Fanuc KAREL source: CA0036.KL

PROGRAM CA0036
%STACKSIZE=65535
%PRIORITY=65535
%NOLOCKGROUP
TYPE
T=STRUCTURE
A : INTEGER
B : REAL
ENDSTRUCTURE
VAR
G : INTEGER
I : INTEGER
R : REAL
B : BOOLEAN
S : STRING[16]
AI : ARRAY[2] OF INTEGER
AR : ARRAY[2] OF REAL
ST : T
P : XYZWPR
V : VECTOR
ROUTINE F(P1 : ARRAY[*] OF INTEGER; P2 : ARRAY[*] OF REAL; P3 : T; P4 : XYZWPR; P5 : VECTOR; P6 : ARRAY[*] OF INTEGER; P7 : ARRAY[*] OF REAL; P8 : T; P9 : XYZWPR; P10 : VECTOR; P11 : ARRAY[*] OF INTEGER;
P12 : ARRAY[*] OF REAL) FROM CA0036
ROUTINE F
BEGIN
G=(G + 1)
END F
BEGIN
G=0
I=1
R=2.5
B=TRUE
S='A'
AI[1]=3
AR[1]=4.5
-- UNSAFE_SOURCE_IR line 42: ST.A = 5
-- UNSAFE_SOURCE_IR line 43: ST.B = 6.5
F(AI,AR,ST,P,V,AI,AR,ST,P,V,AI,AR)
END CA0036
